TYPE ST_ProdParams :
STRUCT
	sTankDescription: STRING;
	arrComponents	: ARRAY [0..g_Prod.cMaxCompInProduct-1] OF ST_Component;
	///Stirrer params
	iStirrerRpm		: UINT;
	iStirrerOnTime	: UINT;
	iStirrerOffTime	: UINT;
	
	//production
	iLitDrainBeforeProd	: UINT;
	rMinTempToStartProd	: REAL;
	rMaxTempToStartProd	: REAL;
	iShelfLife			: UINT;
END_STRUCT
END_TYPE

(* stored: Version 1.1.0.1, ProductVersion 3.1.4024.15
   DUT ST_ProdParams: Id {b0187377-aa66-4e19-a2df-9cc951c4a66e} *)
